// TIA Portal V20 export
// export: Created 2026-10-12T04:58:22.1440736Z, ExportSetting WithDefaults, DisplayName Totally Integrated Automation Portal, DisplayVersion V20, DisplayName TIA Portal Openness, DisplayVersion V20, DisplayName TIA Portal Teamcenter Gateway, DisplayVersion V20, DisplayName TIA Portal Version Control Interface, DisplayVersion V20, DisplayName SINAMICS Startdrive Advanced, DisplayVersion V20 SP1 Update 2, DisplayName SINAMICS Startdrive G110M, G120, G120C, G120D, G120P, G115D, DisplayVersion V20 SP1 Update 2, DisplayName SINAMICS Startdrive G130, G150, S120, S150, SINAMICS MV, G220, S200, S210, DisplayVersion V20 SP1 Update 2, DisplayName STEP 7 Professional, DisplayVersion V20, DisplayName STEP 7 Safety, DisplayVersion V20, DisplayName WinCC Basic/Comfort/Advanced, DisplayVersion V20, DisplayName WinCC Professional, DisplayVersion V20, DisplayName WinCC Unified, DisplayVersion V20
FUNCTION "F_ConfigSetBench" : Void   // FC165, SCL
{ S7_Optimized_Access := 'TRUE' }
VERSION : 0.1
// Test-only tampering: the production retained store stays inaccessible.
// stored: AutoNumber true, IsIECCheckEnabled false, SetENOAutomatically false, UDAEnableTagReadback false
   VAR_TEMP
      Slot : Int;
      Index : Int;
   END_VAR
BEGIN

   IF NOT "GDB_ConfigSetTest".Corrupt THEN
       RETURN;
   END_IF;
   "GDB_ConfigSetTest".Corrupt := FALSE;
   #Slot := "FRK_SetFind"(RootIndex := 1, SetName := "GDB_ConfigSetTest".SetName);
   "GDB_ConfigSetTest".Slot := #Slot;
   IF #Slot = 0 THEN
       RETURN;
   END_IF;
   #Index := "FRK_SetStore".Sets[1, #Slot].Info.RecordCount;
   "GDB_ConfigSetTest".RecordScope := "FRK_SetStore".Sets[1, #Slot].Records[#Index].Scope;
   "GDB_ConfigSetTest".RecordKey := "FRK_SetStore".Sets[1, #Slot].Records[#Index].WriteKey;
   CASE "GDB_ConfigSetTest".Field OF
       1:
           "FRK_SetStore".Sets[1, #Slot].Records[#Index].ValueText := "GDB_ConfigSetTest".Text;
       2:
           "FRK_SetStore".Sets[1, #Slot].Records[#Index].Revision := 99;
       3:
           "FRK_SetStore".Sets[1, #Slot].Records[#Index].ValueType := 99;
       4:
           "FRK_SetStore".Sets[1, #Slot].Records[#Index].WriteKey := 'unknown';
       5:
           "FRK_SetStore".Sets[1, #Slot].Records[#Index].Scope := 'StationB';
       6:
           "FRK_SetStore".Sets[1, #Slot].Info.RecordCount := #Index - 1;
       7:
           "FRK_SetStore".Sets[1, #Slot].Records[#Index] := "FRK_SetStore".Sets[1, #Slot].Records[1];
       ELSE
           RETURN;
   END_CASE;
END_FUNCTION
